KUKA KRL program: FeatureTest.src

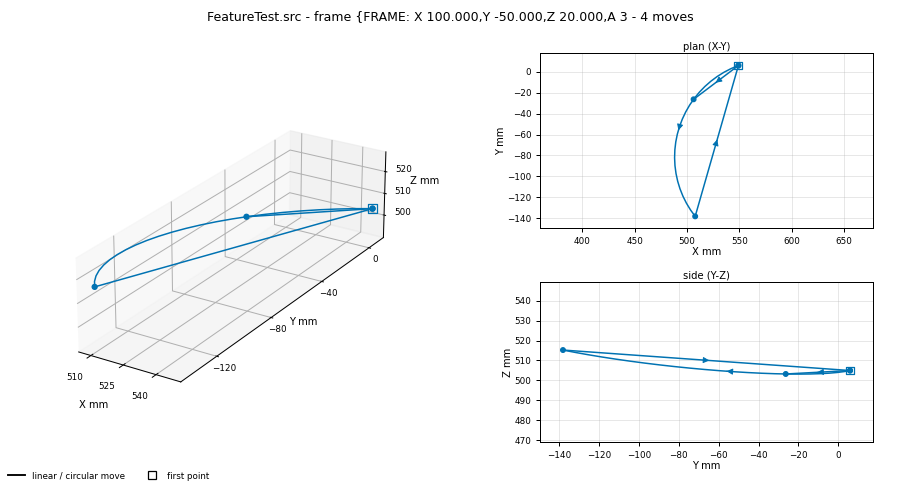
[picture p0: tool path of FeatureTest.src in frame {FRAME: X 100.000,Y -50.000,Z 20.000,A 3, 4 of 6 moves have a stored position in this frame; points joined in program order, loops and branches not executed]
&ACCESS RVP
&REL 1
&PARAM TEMPLATE = C:\KRC\Roboter\Template\vorgabe
&PARAM EDITMASK = *
DEF FeatureTest ( )

; External program calls:
EXT MyFunc()
EXT SetRPM()
EXT SubPick()

EXT BAS (BAS_COMMAND :IN,REAL :IN )


; GLOBAL INTERRUPT DECL 3 WHEN $STOPMESS==TRUE DO IR_STOPM ( )
; INTERRUPT ON 3

;FOLD Initialise and set default speed
BAS (#INITMOV,0)
BAS (#VEL_PTP,100)
BAS (#ACC_PTP,20)
$VEL.CP=0.2
BAS (#TOOL,0)
BAS (#BASE,0)
;ENDFOLD

;;FOLD STARTPOS
;$BWDSTART = FALSE
;PDAT_ACT = PDEFAULT
;BAS(#PTP_DAT)
;FDAT_ACT = {TOOL_NO 0,BASE_NO 0,IPO_FRAME #BASE}
;BAS(#FRAMES)
;;ENDFOLD

$ADVANCE = 5

;FOLD ---- Quickly skip BCO ----
; PTP $AXIS_ACT
;ENDFOLD

;FOLD ---- GO HOME ----
; PTP {A1 0.000, A2 -90.000, A3 90.000, A4 0.000, A5 0.000, A6 0.000, E1 0, E2 0, E3 0, E4 0, E5 0, E6 0}
;ENDFOLD


; Program generated by VerticalBot Studio for KUKA KR 6 R900 sixx on 25/10/2026 12:00:00
; Using nominal kinematics.
; ---- Setting reference (Base) ----
; BASE_DATA[2] = {FRAME: X 100.000,Y -50.000,Z 20.000,A 30.000,B 0.000,C 0.000}
$BASE = {FRAME: X 100.000,Y -50.000,Z 20.000,A 30.000,B 0.000,C 0.000}
; $BASE = BASE_DATA[2]
; --------------------------
; ---- Setting tool (TCP) ----
; TOOL_DATA[1] = {FRAME: X 10.000,Y 0.000,Z 120.000,A 0.000,B 15.000,C 0.000}
$TOOL = {FRAME: X 10.000,Y 0.000,Z 120.000,A 0.000,B 15.000,C 0.000}
; $TOOL = TOOL_DATA[1]
; --------------------------
$VEL.CP = 0.30000
$VEL.ORI1 = 90.00000
$VEL.ORI2 = 90.00000
$ACC.CP = 1.50000
$ACC.ORI1 = 400.00000
$ACC.ORI2 = 400.00000
$APO.CPTP = 5
$APO.CDIS = 5.000
PTP {A1 10.00000,A2 -80.00000,A3 100.00000,A4 20.00000,A5 40.00000,A6 -30.00000} C_PTP
LIN {X 549.094,Y 5.962,Z 504.960,A -174.431,B 15.001,C 175.695} C_DIS
CIRC {X 506.272,Y -26.320,Z 503.226,A -178.509,B 14.048,C 175.384},{X 507.783,Y -138.190,Z 515.247,A 171.653,B 15.955,C 176.009} C_DIS
$VEL.CP = 0.05000
$APO.CPTP = 0
$APO.CDIS = 0.000
LIN {X 549.094,Y 5.962,Z 504.960,A -174.431,B 15.001,C 175.695} C_DIS
$VEL.CP = 0.30000
LIN {X 506.272,Y -26.320,Z 503.226,A -178.509,B 14.048,C 175.384}
$OUT[3]=TRUE
DO_GRIP=FALSE
WAIT FOR ($IN[5]==TRUE)
START_TIMER:
$TIMER_STOP[1]=TRUE
$TIMER_FLAG[1]=FALSE
$TIMER[1]=2.000
$TIMER_STOP[1]=FALSE
WAIT FOR (DI_PART==TRUE OR $TIMER_FLAG[1])
$TIMER_STOP[1]=TRUE
IF $TIMER_FLAG[1]== TRUE THEN
    HALT ; Timed out!
    GOTO START_TIMER
ENDIF
WAIT SEC 0.500
; a comment line
Wait for StrClear($LOOP_MSG[])
$LOOP_CONT = TRUE
$LOOP_MSG[] = "Hello operator"
MyFunc()
SetRPM(5000)
RAW_CODE_LINE
SubPick()
$VEL.ORI1 = 45.00000
$VEL.ORI2 = 45.00000
; ---- Setting tool (TCP) ----
; TOOL_DATA[1] = {FRAME: X 10.000,Y 0.000,Z 120.000,A 0.000,B 15.000,C 0.000}
$TOOL = {FRAME: X 10.000,Y 0.000,Z 120.000,A 0.000,B 15.000,C 0.000}
; $TOOL = TOOL_DATA[1]
; --------------------------
; Attach to Tool 1
PTP {A1 10.00000,A2 -80.00000,A3 100.00000,A4 20.00000,A5 40.00000,A6 -30.00000}
HALT
END
